Fanuc KAREL source: kt00304.KL

-- PROVISIONAL review KL for V770-1; original PC SHA256 37b3b3b92be90ed3983483f8a6a47425c5d903ba70f49ed784cfac004115d6ab
-- Incomplete behavior may be omitted. Consult companion uncertainty JSON. Do not deploy.
PROGRAM KT00304
%NOLOCKGROUP
VAR
  R2 : REAL
  OUT : BOOLEAN
-- UNRESOLVED_DECL Y1 type=002018
BEGIN
  -- UNRESOLVED_PC offsets 5-19; opcodes 2E,22,9D,33,B2
  -- UNRESOLVED_PC offsets 24-35; opcodes 2E,23
  -- UNRESOLVED_PC offsets 40-64; opcodes 22,9D,33,B1,21,29,64,6E,23
  -- UNRESOLVED_PC offsets 69-73; opcodes 7F
END KT00304
